PROGRAM ExampleProgram2
VAR
	fbTimerOff  : TON;
    fbTimerOn   : TON;
    tOffTime    : TIME := T#1000MS; // Mappable off-time
    tOnTime     : TIME := T#1000MS; // Mappable on-time
    bBlinkerOn  : BOOL;
	bBlinkerOff : BOOL;
END_VAR

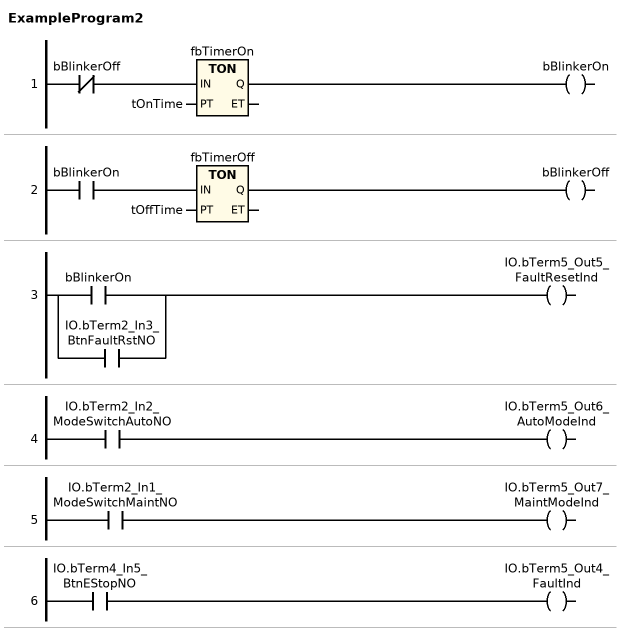
// NETWORK 1
fbTimerOn(IN := NOT bBlinkerOff, PT := tOnTime); // TON
bBlinkerOn := fbTimerOn.Q;

// NETWORK 2
fbTimerOff(IN := bBlinkerOn, PT := tOffTime); // TON
bBlinkerOff := fbTimerOff.Q;

// NETWORK 3
IO.bTerm5_Out5_FaultResetInd := bBlinkerOn OR IO.bTerm2_In3_BtnFaultRstNO;

// NETWORK 4
IO.bTerm5_Out6_AutoModeInd := IO.bTerm2_In2_ModeSwitchAutoNO;

// NETWORK 5
IO.bTerm5_Out7_MaintModeInd := IO.bTerm2_In1_ModeSwitchMaintNO;

// NETWORK 6
IO.bTerm5_Out4_FaultInd := IO.bTerm4_In5_BtnEStopNO;

END_PROGRAM

(* stored: Version 1.1.0.1, ProductVersion 3.1.4024.16
   POU ExampleProgram2: Id {7cf0928f-9d39-4b48-8542-e2949f969e22}, SpecialFunc None *)
